FUNCTION_BLOCK FB_TriBlender_Select EXTENDS FB_SFC_Cycle IMPLEMENTS ITF_FB_SFC_Cycle
VAR_INPUT
	valInSelect		: E_Pis_Name;
	valInMarinade	: E_Pis_Name;
	valInColor		: E_Pis_Name;
	valOutSelect	: E_Pis_Name;	
	valOutMarinade	: E_Pis_Name;
	valOutColor		: E_Pis_Name;
	valDrain		: E_Pis_Name;
	
END_VAR
VAR_OUTPUT
END_VAR
VAR
	//refElement		: REFERENCE TO FB_Element;
	//refState_Long		: REFERENCE TO E_Element_State_Long;
	eReq				: E_TriBlenderSelect;
	eProcess			: E_TriBlenderSelect;
	eStatus				: E_TriBlenderSelect;
	
	fbPis				: FB_Piston;
	stPis_InSelect		: REFERENCE TO ST_Piston;
	stPis_InMarinade	: REFERENCE TO ST_Piston;
	stPis_InColor		: REFERENCE TO ST_Piston;
	stPis_OutSelect		: REFERENCE TO ST_Piston;
	stPis_OutMarinade	: REFERENCE TO ST_Piston;
	stPis_OutColor		: REFERENCE TO ST_Piston;
	stPis_Drain			: REFERENCE TO ST_Piston;

	tonDrainTime: TON;
	rt_Req_Reset: R_TRIG;
	//bRun: BOOL;
	//bDone: BOOL;
	SFCReset: BOOL;
	//bStepDone: BOOL;
END_VAR
VAR_IN_OUT


END_VAR

act_GetReference();

act_Oper();
IF NOT Init.x THEN;
	act_Status();
END_IF

tonDrainTime(PT:=T#1M, IN:=eStatus=E_TriBlenderSelect.eDrain);
IF tonDrainTime.Q 
AND eReq=E_TriBlenderSelect.eNone
AND eProcess=E_TriBlenderSelect.eNone
THEN;
	eReq:=E_TriBlenderSelect.eMarinade;
END_IF

m_Request_Reset(memo:=rt_Req_Reset);//

ACTION _aColor_1_active:
bStepDone:=FALSE;
IF TRUE 
AND eStatus=E_TriBlenderSelect.eColor
THEN;
	bStepDone:=TRUE;
END_IF
END_ACTION

ACTION _aColor_1_entry:
fbPis.m_SetByRecipe(stPis:=stPis_InSelect, 			req:=E_Piston_Recipe_State.Act);
fbPis.m_SetByRecipe(stPis:=stPis_InMarinade, 		req:=E_Piston_Recipe_State.Release);
fbPis.m_SetByRecipe(stPis:=stPis_InColor, 			req:=E_Piston_Recipe_State.Release);
fbPis.m_SetByRecipe(stPis:=stPis_OutSelect, 		req:=E_Piston_Recipe_State.Act);
fbPis.m_SetByRecipe(stPis:=stPis_OutMarinade, 		req:=E_Piston_Recipe_State.Release);
fbPis.m_SetByRecipe(stPis:=stPis_OutColor, 			req:=E_Piston_Recipe_State.Release);
fbPis.m_SetByRecipe(stPis:=stPis_Drain, 			req:=E_Piston_Recipe_State.Release);
END_ACTION

ACTION _aColor_2_entry:
fbPis.m_SetByRecipe(stPis:=stPis_Drain, 			req:=E_Piston_Recipe_State.Act);
END_ACTION

ACTION _aColor_3_active:
bStepDone:=FALSE;
IF TRUE 
AND eStatus=E_TriBlenderSelect.eColor
THEN;
	bStepDone:=TRUE;
END_IF
END_ACTION

ACTION _aColor_3_entry:
fbPis.m_SetByRecipe(stPis:=stPis_InSelect, 			req:=E_Piston_Recipe_State.Act);
fbPis.m_SetByRecipe(stPis:=stPis_InMarinade, 		req:=E_Piston_Recipe_State.Release);
fbPis.m_SetByRecipe(stPis:=stPis_InColor, 			req:=E_Piston_Recipe_State.Release);
fbPis.m_SetByRecipe(stPis:=stPis_OutSelect, 		req:=E_Piston_Recipe_State.Act);
fbPis.m_SetByRecipe(stPis:=stPis_OutMarinade, 		req:=E_Piston_Recipe_State.Release);
fbPis.m_SetByRecipe(stPis:=stPis_OutColor, 			req:=E_Piston_Recipe_State.Release);
fbPis.m_SetByRecipe(stPis:=stPis_Drain, 			req:=E_Piston_Recipe_State.Release);
END_ACTION

ACTION _aDone_entry:
eProcess:=E_TriBlenderSelect.eNone;
eReq:=E_TriBlenderSelect.eNone;
eStatus:=E_TriBlenderSelect.eNone;
bRun:=FALSE;
bDone:=TRUE;
END_ACTION

ACTION _aDrain_active:
bStepDone:=FALSE;
IF TRUE 
AND eStatus=E_TriBlenderSelect.eDrain
THEN;
	bStepDone:=TRUE;
END_IF
END_ACTION

ACTION _aDrain_entry:
fbPis.m_SetByRecipe(stPis:=stPis_InSelect, 			req:=E_Piston_Recipe_State.Release);
fbPis.m_SetByRecipe(stPis:=stPis_InMarinade, 		req:=E_Piston_Recipe_State.Act);
fbPis.m_SetByRecipe(stPis:=stPis_InColor, 			req:=E_Piston_Recipe_State.Act);
fbPis.m_SetByRecipe(stPis:=stPis_OutSelect, 		req:=E_Piston_Recipe_State.Release);
fbPis.m_SetByRecipe(stPis:=stPis_OutMarinade, 		req:=E_Piston_Recipe_State.Act);
fbPis.m_SetByRecipe(stPis:=stPis_OutColor, 			req:=E_Piston_Recipe_State.Act);
fbPis.m_SetByRecipe(stPis:=stPis_Drain, 			req:=E_Piston_Recipe_State.Act);
END_ACTION

ACTION _aInit_active:
SFCReset:=FALSE;
END_ACTION

ACTION _aMarinade_1_active:
bStepDone:=FALSE;
IF TRUE 
AND eStatus=E_TriBlenderSelect.eMarinade
THEN;
	bStepDone:=TRUE;
END_IF
END_ACTION

ACTION _aMarinade_1_entry:
fbPis.m_SetByRecipe(stPis:=stPis_InSelect, 			req:=E_Piston_Recipe_State.Release);
fbPis.m_SetByRecipe(stPis:=stPis_InMarinade, 		req:=E_Piston_Recipe_State.Release);
fbPis.m_SetByRecipe(stPis:=stPis_InColor, 			req:=E_Piston_Recipe_State.Release);
fbPis.m_SetByRecipe(stPis:=stPis_OutSelect, 		req:=E_Piston_Recipe_State.Release);
fbPis.m_SetByRecipe(stPis:=stPis_OutMarinade, 		req:=E_Piston_Recipe_State.Release);
fbPis.m_SetByRecipe(stPis:=stPis_OutColor, 			req:=E_Piston_Recipe_State.Release);
fbPis.m_SetByRecipe(stPis:=stPis_Drain, 			req:=E_Piston_Recipe_State.Release);
END_ACTION

ACTION _aMarinade_2_entry:
fbPis.m_SetByRecipe(stPis:=stPis_Drain, 			req:=E_Piston_Recipe_State.Act);
END_ACTION

ACTION _aMarinade_3_active:
bStepDone:=FALSE;
IF TRUE 
AND eStatus=E_TriBlenderSelect.eMarinade
THEN;
	bStepDone:=TRUE;
END_IF
END_ACTION

ACTION _aMarinade_3_entry:
fbPis.m_SetByRecipe(stPis:=stPis_InSelect, 			req:=E_Piston_Recipe_State.Release);
fbPis.m_SetByRecipe(stPis:=stPis_InMarinade, 		req:=E_Piston_Recipe_State.Release);
fbPis.m_SetByRecipe(stPis:=stPis_InColor, 			req:=E_Piston_Recipe_State.Release);
fbPis.m_SetByRecipe(stPis:=stPis_OutSelect, 		req:=E_Piston_Recipe_State.Release);
fbPis.m_SetByRecipe(stPis:=stPis_OutMarinade, 		req:=E_Piston_Recipe_State.Release);
fbPis.m_SetByRecipe(stPis:=stPis_OutColor, 			req:=E_Piston_Recipe_State.Release);
fbPis.m_SetByRecipe(stPis:=stPis_Drain, 			req:=E_Piston_Recipe_State.Release);
END_ACTION

ACTION _aReady_active:

eStatus:=E_TriBlenderSelect.eNone;
CASE eReq OF
	E_TriBlenderSelect.eColor:;
			IF TRUE THEN;
				eProcess:=E_TriBlenderSelect.eColor;
			END_IF	
			
	E_TriBlenderSelect.eDrain:;
			IF TRUE THEN;
				eProcess:=E_TriBlenderSelect.eDrain;
			END_IF
			
	E_TriBlenderSelect.eMarinade:;
			IF TRUE THEN;
				eProcess:=E_TriBlenderSelect.eMarinade;
			END_IF

END_CASE
END_ACTION

ACTION act_GetReference:
m_Set_SFCFlags_Reference();
//refElement REF= fbElement[eElementID];

stPis_InSelect	 REF= g_Piston.stPis[valInSelect];
stPis_InMarinade REF= g_Piston.stPis[valInMarinade];
stPis_InColor	 REF= g_Piston.stPis[valInColor];

stPis_OutSelect	  REF= g_Piston.stPis[valOutSelect];
stPis_OutMarinade REF= g_Piston.stPis[valOutMarinade];
stPis_OutColor	  REF= g_Piston.stPis[valOutColor];

stPis_Drain		  REF= g_Piston.stPis[valDrain];
END_ACTION

ACTION act_Oper:
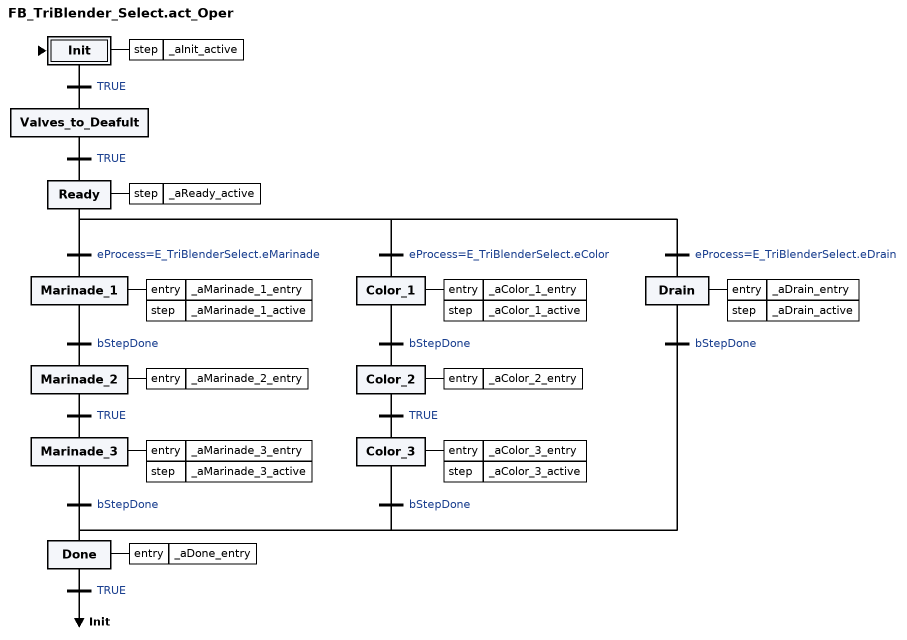
INITIAL_STEP Init:
    _aInit_active(N);  // step action
END_STEP
TRANSITION FROM Init TO Valves_to_Deafult
    := TRUE;
END_TRANSITION
STEP Valves_to_Deafult:
END_STEP
TRANSITION FROM Valves_to_Deafult TO Ready
    := TRUE;
END_TRANSITION
STEP Ready:
    _aReady_active(N);  // step action
END_STEP
TRANSITION FROM Ready TO Marinade_1
    := eProcess=E_TriBlenderSelect.eMarinade;
END_TRANSITION
STEP Marinade_1:
    _aMarinade_1_entry(P1);  // entry action
    _aMarinade_1_active(N);  // step action
END_STEP
TRANSITION FROM Marinade_1 TO Marinade_2
    := bStepDone;
END_TRANSITION
STEP Marinade_2:  // min time T#10s
    _aMarinade_2_entry(P1);  // entry action
END_STEP
TRANSITION FROM Marinade_2 TO Marinade_3
    := TRUE;
END_TRANSITION
STEP Marinade_3:
    _aMarinade_3_entry(P1);  // entry action
    _aMarinade_3_active(N);  // step action
END_STEP
TRANSITION FROM Marinade_3 TO Done
    := bStepDone;
END_TRANSITION
TRANSITION FROM Ready TO Color_1
    := eProcess=E_TriBlenderSelect.eColor;
END_TRANSITION
STEP Color_1:
    _aColor_1_entry(P1);  // entry action
    _aColor_1_active(N);  // step action
END_STEP
TRANSITION FROM Color_1 TO Color_2
    := bStepDone;
END_TRANSITION
STEP Color_2:  // min time T#10s
    _aColor_2_entry(P1);  // entry action
END_STEP
TRANSITION FROM Color_2 TO Color_3
    := TRUE;
END_TRANSITION
STEP Color_3:
    _aColor_3_entry(P1);  // entry action
    _aColor_3_active(N);  // step action
END_STEP
TRANSITION FROM Color_3 TO Done
    := bStepDone;
END_TRANSITION
TRANSITION FROM Ready TO Drain
    := eProcess=E_TriBlenderSelect.eDrain;
END_TRANSITION
STEP Drain:
    _aDrain_entry(P1);  // entry action
    _aDrain_active(N);  // step action
END_STEP
TRANSITION FROM Drain TO Done
    := bStepDone;
END_TRANSITION
STEP Done:  // min time T#0.2s
    _aDone_entry(P1);  // entry action
END_STEP
TRANSITION FROM Done TO Init
    := TRUE;
END_TRANSITION
// branch label Branch0_act_Oper_Tank
END_ACTION

ACTION act_Status:
IF TRUE 
AND fbPis.m_CheckByRecipe(stPis:=stPis_InSelect, 		req:=E_Piston_Recipe_State.Release)
AND fbPis.m_CheckByRecipe(stPis:=stPis_InMarinade, 		req:=E_Piston_Recipe_State.Release)
AND fbPis.m_CheckByRecipe(stPis:=stPis_InColor, 		req:=E_Piston_Recipe_State.Release)
AND fbPis.m_CheckByRecipe(stPis:=stPis_OutSelect, 		req:=E_Piston_Recipe_State.Release)
AND fbPis.m_CheckByRecipe(stPis:=stPis_OutMarinade, 	req:=E_Piston_Recipe_State.Release)
AND fbPis.m_CheckByRecipe(stPis:=stPis_OutColor, 		req:=E_Piston_Recipe_State.Release)
AND fbPis.m_CheckByRecipe(stPis:=stPis_Drain	, 		req:=E_Piston_Recipe_State.Release)
THEN;
	eStatus:=E_TriBlenderSelect.eMarinade;
	
ELSIF TRUE 
AND fbPis.m_CheckByRecipe(stPis:=stPis_InSelect, 		req:=E_Piston_Recipe_State.Act)
AND fbPis.m_CheckByRecipe(stPis:=stPis_InMarinade, 		req:=E_Piston_Recipe_State.Release)
AND fbPis.m_CheckByRecipe(stPis:=stPis_InColor, 		req:=E_Piston_Recipe_State.Release)
AND fbPis.m_CheckByRecipe(stPis:=stPis_OutSelect, 		req:=E_Piston_Recipe_State.Act)
AND fbPis.m_CheckByRecipe(stPis:=stPis_OutMarinade, 	req:=E_Piston_Recipe_State.Release)
AND fbPis.m_CheckByRecipe(stPis:=stPis_OutColor, 		req:=E_Piston_Recipe_State.Release)
AND fbPis.m_CheckByRecipe(stPis:=stPis_Drain	, 		req:=E_Piston_Recipe_State.Release)
THEN;
	eStatus:=E_TriBlenderSelect.eColor;
	
ELSIF TRUE 
AND fbPis.m_CheckByRecipe(stPis:=stPis_InSelect, 		req:=E_Piston_Recipe_State.Release)
AND fbPis.m_CheckByRecipe(stPis:=stPis_InMarinade, 		req:=E_Piston_Recipe_State.Act)
AND fbPis.m_CheckByRecipe(stPis:=stPis_InColor, 		req:=E_Piston_Recipe_State.Act)
AND fbPis.m_CheckByRecipe(stPis:=stPis_OutSelect, 		req:=E_Piston_Recipe_State.Release)
AND fbPis.m_CheckByRecipe(stPis:=stPis_OutMarinade, 	req:=E_Piston_Recipe_State.Act)
AND fbPis.m_CheckByRecipe(stPis:=stPis_OutColor, 		req:=E_Piston_Recipe_State.Act)
AND fbPis.m_CheckByRecipe(stPis:=stPis_Drain	, 		req:=E_Piston_Recipe_State.Act)
THEN;
	eStatus:=E_TriBlenderSelect.eDrain;
	
ELSE
	eStatus:=E_TriBlenderSelect.eNone;
	
END_IF;
END_ACTION

METHOD m_CheckStatus : BOOL
VAR_INPUT
	eReqStatus		: E_TriBlenderSelect;
END_VAR
IF eStatus=eReqStatus 
AND eProcess=E_TriBlenderSelect.eNone
AND eReq=E_TriBlenderSelect.eNone
AND bReady
AND bDone
AND NOT bRun
THEN;
	m_CheckStatus:=TRUE;
END_IF
END_METHOD

METHOD m_Request_Reset : BOOL
VAR_IN_OUT
	memo: R_TRIG;
END_VAR
memo(CLK:=eReq=0);
IF TRUE 
AND memo.Q
THEN;
	SFCReset:=TRUE;
END_IF
END_METHOD

METHOD m_Run : BOOL
VAR_INPUT
	eReqProc			: E_TriBlenderSelect;
END_VAR
IF eProcess=E_TriBlenderSelect.eNone THEN;
	eProcess:=eReq:=eReqProc;
	bDone:=FALSE;
	m_Run:=TRUE;
END_IF
END_METHOD

METHOD m_Set_Request : BOOL
VAR_INPUT
	eSetReg		: E_TriBlenderSelect;
END_VAR
eReq:=eSetReg;
END_METHOD

{warning 'add method implementation '}
METHOD m_Set_SFCFlags_Reference : BOOL
//Set reference to SFC flags

refSFC.SFCInit REF= SFCInit;
refSFC.SFCReset REF= SFCReset;
refSFC.SFCError REF= SFCError;
refSFC.SFCEnableLimit REF= SFCEnableLimit;
refSFC.SFCErrorStep REF= SFCErrorStep;
refSFC.SFCErrorPOU REF= SFCErrorPOU;
refSFC.SFCQuitError REF= SFCQuitError;
refSFC.SFCPause REF= SFCPause;
refSFC.SFCTrans REF= SFCTrans;
refSFC.SFCCurrentStep REF= SFCCurrentStep;
refSFC.SFCTip REF= SFCTip;
refSFC.SFCTipMode REF= SFCTipMode;

// Cycle handle for SFC
m_SFC_Handle();
END_METHOD

END_FUNCTION_BLOCK

(* stored: Version 1.1.0.1, ProductVersion 3.1.4024.15
   POU FB_TriBlender_Select: Id {9eeca8ec-03ab-4735-83e4-c97ea5515e09}, SpecialFunc None
   Folder Manage: Id {e20a7cbd-7252-4410-8f32-fdf6c8d5cc66}
   Action _aColor_1_active: Id {0e00c0e9-109c-44f6-b8b4-7e71627c84d3}
   Action _aColor_1_entry: Id {b8924bfb-9851-4d09-8b08-65fd1d78ee0f}
   Action _aColor_2_entry: Id {da1ef349-ea15-4f48-b15c-f9a0538473e0}
   Action _aColor_3_active: Id {03ef5e54-1af1-417a-ae7a-2b87b7ca015f}
   Action _aColor_3_entry: Id {d09ad859-038c-4689-aa9b-288e4360d209}
   Action _aDone_entry: Id {cb123ed7-cd01-4641-ac5c-2e5e006fc25a}
   Action _aDrain_active: Id {96576044-f427-44d6-9d13-e5ce72838ebe}
   Action _aDrain_entry: Id {7d00fb3f-348c-4f15-b27d-345a85d5f604}
   Action _aInit_active: Id {6a7b3ace-94ba-4ea9-b6fb-bb0533f3c28a}
   Action _aMarinade_1_active: Id {82658e7b-8830-47dc-acf2-53cf20863f1a}
   Action _aMarinade_1_entry: Id {ba08c11b-233b-4723-8599-c0e89d2ffeb8}
   Action _aMarinade_2_entry: Id {5ff3c56b-3111-449c-a5be-278c24186f0e}
   Action _aMarinade_3_active: Id {c5b58539-e354-46aa-9ffb-6ea148a749e2}
   Action _aMarinade_3_entry: Id {85ef1959-4baa-48bf-ba34-61599ccb810d}
   Action _aReady_active: Id {e9c65ea6-1cf6-4665-b228-f295655c142c}
   Action act_GetReference: Id {1f7e6d9f-c733-467c-bd8d-99c3278d05fb}
   Action act_Oper: Id {b80f5ade-5ea6-4341-a41a-f2c6d43c3182}
   Action act_Status: Id {09075606-aba2-4421-aadf-8a8f6410b267}
   Method m_CheckStatus: Id {3903e6c5-5909-4217-872b-04f94cc50c95}
   Method m_Request_Reset: Id {6dfb826e-0c5a-4b01-8291-56a11557903f}
   Method m_Run: Id {a8b44bf2-fd16-4b21-9c83-6e8184bbb941}
   Method m_Set_Request: Id {a1fa741f-11b0-4781-a2c4-c8fa2ef789ea}
   Method m_Set_SFCFlags_Reference: Id {40d7e9fd-d4fa-45bd-88e4-d85c0e80f0bc} *)
